// TIA Portal V21 export
ORGANIZATION_BLOCK "Series"   // OB1, LAD
BEGIN

REGION Network 1: Motor run
   // Start, unless stopped.
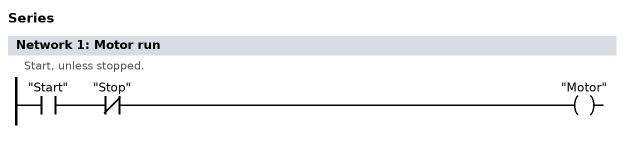
   RUNG wire#powerrail
      Contact( "Start" )
      I_Contact( "Stop" )
      Coil( "Motor" )
   END_RUNG
   // the same network as SCL:
   "Motor" := "Start" AND NOT "Stop";
END_REGION
END_ORGANIZATION_BLOCK
